FUNCTION_BLOCK FB_MotorFake EXTENDS FB_MotorBase
VAR_INPUT
    fault : BOOL;
END_VAR

SUPER^();

METHOD PROTECTED CheckFault : BOOL
(* SUPER selects the base hook, while inherited Update dispatches here. *)
CheckFault := SUPER^.CheckFault() OR fault;
END_METHOD

END_FUNCTION_BLOCK

(* stored: Version 1.1.0.1, ProductVersion 3.1 *)
